// On-delay timer for the long command timeouts. Same behaviour as TON, but the preset time is divided by nDivisor
// (default 1), so a test can run a 12 h timeout in a few scans. The divisor is an input of the owner (per instance, not
// a global): TcUnit runs all suites in the same PLC cycles, so a global would shorten the timeouts of every running test.
FUNCTION_BLOCK FB_TimeoutTimer
VAR_INPUT
	IN	: BOOL;
	PT	: TIME;
	nDivisor	: UDINT := 1;
END_VAR
VAR_OUTPUT
	Q	: BOOL;
	ET	: TIME;
END_VAR
VAR
	ton	: TON;
END_VAR

IF nDivisor > 1 THEN
	ton(IN := IN, PT := DWORD_TO_TIME(TIME_TO_DWORD(PT) / nDivisor), Q => Q, ET => ET);
ELSE
	ton(IN := IN, PT := PT, Q => Q, ET => ET);
END_IF

END_FUNCTION_BLOCK

(* stored: Version 1.1.0.1, ProductVersion 3.1.4024.15
   POU FB_TimeoutTimer: Id {be2effaf-8032-44f0-b85c-850071e4590c}, SpecialFunc None *)
